// TIA Portal V21 export
Screen "T08_Bar"  1024x768, Number=28
  ScreenLayer 
    Bar "P_Bar" at 0,0 size 100x30  MaximumValue=24
      ProcessValue := BalL
